// TIA Portal V21 export
// export: Created 2026-11-10T23:32:28.9908613Z, ExportSetting WithDefaults, DisplayName Totally Integrated Automation Portal, DisplayVersion V21 Update 3, DisplayName STEP 7 Professional, DisplayVersion V21 Update 3, DisplayName STEP 7 Safety, DisplayVersion V21, DisplayName Tech WebApplication, DisplayVersion V21, DisplayName WinCC Basic/Comfort/Advanced, DisplayVersion V21 Update 3, DisplayName WinCC Unified, DisplayVersion V21 Update 3
DATA_BLOCK "mTO_ExternalEncoder"   // DB8, Motion_DB
// stored: AutoNumber true, DBAccessibleFromOPCUA true, DBAccessibleFromWebserver true, InstanceOfName TO_ExternalEncoder, OfSystemLibElement TO_ExternalEncoder, OfSystemLibVersion 8.0
TO_ExternalEncoder   // technology object, version 8.0
// stored: Connection Interface Sensor, SensorIndexInActorTelegram 1, PathToDBMember DB_Enc.tel.Sensor_1
   // // inherited from TO_Axis
   // // inherited from TO_Object
   // VAR
   //    ActualPosition { ExternalWritable := 'False'} : LReal;
   //    ActualVelocity { ExternalWritable := 'False'} : LReal;
   //    ActualAcceleration { ExternalWritable := 'False'} : LReal;
   //    ActualModuloCycle { ExternalWritable := 'False'} : DInt;
   //    Sensor { S7_SetPoint := 'True'} : TO_Struct_ExternalEncoder_Sensor;
   //    CrossPlcSynchronousOperation { S7_SetPoint := 'True'} : TO_Struct_CrossPlcSynchronousOperation;
   //    Extrapolation { S7_SetPoint := 'True'} : TO_Struct_Extrapolation;
   //    Mechanics { S7_SetPoint := 'True'} : TO_Struct_Mechanics;
   //    LoadGear { S7_SetPoint := 'True'} : TO_Struct_LoadGear;
   //    Properties { ExternalWritable := 'False'; S7_SetPoint := 'True'} : TO_Struct_Properties;
   //    Modulo { S7_SetPoint := 'True'} : TO_Struct_Modulo;
   //    Homing { S7_SetPoint := 'True'} : TO_Struct_ExternalEncoder_Homing;
   //    StandstillSignal { S7_SetPoint := 'True'} : TO_Struct_StandstillSignal;
   //    Units { ExternalWritable := 'False'; S7_SetPoint := 'True'} : TO_Struct_ExternalEncoder_Units;
   //    StatusProvidedLeadingValue { ExternalWritable := 'False'; S7_SetPoint := 'True'} : TO_Struct_StatusProvidedLeadingValue;
   //    StatusSensor { ExternalWritable := 'False'; S7_SetPoint := 'True'} : TO_Struct_StatusSensor;
   //    StatusExtrapolation { ExternalWritable := 'False'; S7_SetPoint := 'True'} : TO_Struct_StatusExtrapolation;
   //    StatusWord { ExternalWritable := 'False'} : DWord;
   //    ErrorWord { ExternalWritable := 'False'} : DWord;
   //    ErrorDetail { ExternalWritable := 'False'; S7_SetPoint := 'True'} : TO_Struct_ErrorDetail;
   //    WarningWord { ExternalWritable := 'False'} : DWord;
   //    InternalToTrace { S7_SetPoint := 'True'} : Array[1..4] of TO_Struct_Internal;
   // END_VAR
BEGIN
   Sensor.Interface.AddressIn.RID := 16#208070e;
   Sensor.Interface.AddressIn.AREA := 16#84;
   Sensor.Interface.AddressIn.DB_NUMBER := 15;
   Sensor.Interface.AddressOut.RID := 16#208070f;
   Sensor.Interface.AddressOut.AREA := 16#84;
   Sensor.Interface.AddressOut.DB_NUMBER := 15;
   Sensor.Interface.AddressOut.OFFSET := 96;
   _Sensor.Interface.Telegram := 81;
END_DATA_BLOCK
